TYPE ST_DosingProcessSimStatus :
STRUCT
	mainFlow			: LREAL; //simulated main flow in l/min
	dosingFlow			: LREAL; //simulated dosing flow in l/min
END_STRUCT
END_TYPE

(* stored: Version 1.1.0.1, ProductVersion 3.1.4024.12
   DUT ST_DosingProcessSimStatus: Id {19e1d628-a713-405d-afcc-00f5ea61afd1} *)
